FUNCTION_BLOCK MotorControl_AOI (* Migrated from Rockwell AOI *)
  (* Standard: 61499-2 *)
  (* Version 1.0, 2026-11-06, st2fb *)
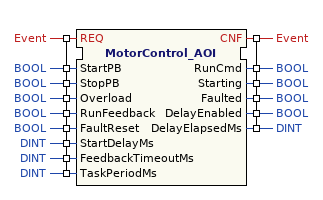
  EVENT_INPUT
    REQ WITH StartPB, StopPB, Overload, RunFeedback, FaultReset, StartDelayMs, FeedbackTimeoutMs, TaskPeriodMs;
  END_EVENT
  EVENT_OUTPUT
    CNF WITH RunCmd, Starting, Faulted, DelayEnabled, DelayElapsedMs;
  END_EVENT
  VAR_INPUT
    StartPB : BOOL;
    StopPB : BOOL;
    Overload : BOOL;
    RunFeedback : BOOL;
    FaultReset : BOOL;
    StartDelayMs : DINT;
    FeedbackTimeoutMs : DINT;
    TaskPeriodMs : DINT;
  END_VAR
  VAR_OUTPUT
    RunCmd : BOOL;
    Starting : BOOL;
    Faulted : BOOL;
    DelayEnabled : BOOL;
    DelayElapsedMs : DINT;
  END_VAR
  VAR
    SD_EN : BOOL := FALSE;
    SD_TT : BOOL := FALSE;
    SD_DN : BOOL := FALSE;
    SD_ACC : DINT := 0;
    SD_PRE : DINT := 0;
    SD_PREV : BOOL := FALSE;
    FT_EN : BOOL := FALSE;
    FT_TT : BOOL := FALSE;
    FT_DN : BOOL := FALSE;
    FT_ACC : DINT := 0;
    FT_PRE : DINT := 0;
    FT_PREV : BOOL := FALSE;
    OS_PREV : BOOL := FALSE;
    OS_OUT : BOOL := FALSE;
    RunLatch : BOOL := FALSE;
    FaultLatch : BOOL := FALSE;
  END_VAR
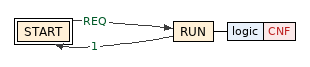
  EC_STATES
    START;
    RUN : logic -> CNF;
  END_STATES
  EC_TRANSITIONS
    START TO RUN := REQ;
    RUN TO START := 1;
  END_TRANSITIONS
  ALGORITHM logic IN ST:
OS_OUT := StartPB AND NOT OS_PREV;
OS_PREV := StartPB;

IF StopPB OR Overload OR FaultLatch THEN
  RunLatch := FALSE;
ELSIF OS_OUT THEN
  RunLatch := TRUE;
END_IF;

SD_EN := RunLatch;
SD_PRE := StartDelayMs;
IF SD_EN THEN
  IF SD_PREV AND NOT SD_DN THEN
    SD_ACC := SD_ACC + TaskPeriodMs;
    IF SD_ACC >= SD_PRE THEN
      SD_ACC := SD_PRE;
      SD_DN := TRUE;
    END_IF;
  END_IF;
ELSE
  SD_ACC := 0;
  SD_DN := FALSE;
END_IF;
SD_TT := SD_EN AND NOT SD_DN;
SD_PREV := SD_EN;
Starting := SD_TT;
RunCmd := SD_DN;
DelayEnabled := SD_EN;
DelayElapsedMs := SD_ACC;

FT_EN := RunCmd AND NOT RunFeedback;
FT_PRE := FeedbackTimeoutMs;
IF FT_EN THEN
  IF FT_PREV AND NOT FT_DN THEN
    FT_ACC := FT_ACC + TaskPeriodMs;
    IF FT_ACC >= FT_PRE THEN
      FT_ACC := FT_PRE;
      FT_DN := TRUE;
    END_IF;
  END_IF;
ELSE
  FT_ACC := 0;
  FT_DN := FALSE;
END_IF;
FT_TT := FT_EN AND NOT FT_DN;
FT_PREV := FT_EN;

IF FT_DN OR Overload THEN
  FaultLatch := TRUE;
END_IF;
IF FaultReset AND NOT Overload THEN
  FaultLatch := FALSE;
  FT_ACC := 0;
  FT_EN := FALSE;
  FT_TT := FALSE;
  FT_DN := FALSE;
  FT_PREV := FALSE;
END_IF;
Faulted := FaultLatch;
  END_ALGORITHM
END_FUNCTION_BLOCK
